Fanuc KAREL source: IO0199.KL

PROGRAM IO0199
%NOLOCKGROUP
%ENVIRONMENT REGOPE
ROUTINE RTEST
VAR
  I : INTEGER
  STATUS : INTEGER
  ENTRY : INTEGER
  A : ARRAY[3] OF INTEGER
  B : BOOLEAN
  R : REAL
  P : XYZWPR
  JPOS : JOINTPOS
  PF : POSITION
BEGIN
  I = 1
  A[1] = 2
  B = TRUE
  R = 1.0
  JPOS = GET_JPOS_REG(1,STATUS,1)
END RTEST
BEGIN
  RTEST
END IO0199
